Fanuc KAREL source: kt00580.compact.KL

PROGRAM KT00580
%STACKSIZE=65535
%PRIORITY=65535
%NOLOCKGROUP
VAR
V1 : VECTOR
I2 : INTEGER
OUT : VECTOR
BEGIN
V1.X=1.0
I2=3
OUT=(V1 / I2)
END KT00580
